// #279: FB_NullComm that records every PublishLog message (not the publishes) in call order. Up to 16; more are counted in
// nOverflow. Clear() empties it. #287: every message that contains sWatch (not empty) is counted in nWatchHits, also past 16.
FUNCTION_BLOCK FB_LogRecordingComm EXTENDS FB_NullComm
VAR_INPUT
	sWatch		: STRING(80);
END_VAR
VAR_OUTPUT
	nWatchHits	: INT;
	nCount		: INT;
	nOverflow	: INT;
	aMessage	: ARRAY[1..16] OF STRING(80);
END_VAR

METHOD Clear
VAR
	i	: INT;
END_VAR
nCount := 0;
nOverflow := 0;
nWatchHits := 0;
FOR i := 1 TO 16 DO
	aMessage[i] := '';
END_FOR
END_METHOD

METHOD PublishLog : BOOL
VAR_INPUT
	level		: STRING(255) := 'INFO';
	message		: STRING(255);
END_VAR
VAR_OUTPUT
	published	: BOOL;
END_VAR
IF LEN(sWatch) > 0 AND FIND(message, sWatch) > 0 THEN
	nWatchHits := nWatchHits + 1;
END_IF
IF nCount >= 16 THEN
	nOverflow := nOverflow + 1;
ELSE
	nCount := nCount + 1;
	aMessage[nCount] := message;
END_IF
PublishLog := TRUE;
published := TRUE;
END_METHOD

END_FUNCTION_BLOCK

(* stored: Version 1.1.0.1, ProductVersion 3.1.4024.15
   POU FB_LogRecordingComm: Id {3857259c-964c-496b-8e74-26e6acc63b48}, SpecialFunc None
   Method Clear: Id {3ec2c5ea-d07f-433c-8fb0-5abd4aeb2cb6}
   Method PublishLog: Id {8f409ef7-e131-4a9f-b1e3-f808f2d8ce69} *)
